(* IEC 61131-3 sources: codesys-to-astra/cds2astra/tests/corpus/C2A-LANG-OOP/pos/src/POUs/FB_B, 1 file *)

(* ---- FB_B.decl.st ---- *)
// Назначение: корпус правила cds2astra (synthetic).
// Автор:      kr0nsch
// Версия:     0.1.0
// Документ:   docs/RULES.md
FUNCTION_BLOCK FB_B EXTENDS FB_A
VAR
END_VAR
